TYPE ST_PolarIIChamber_HolderServiceCtrl :
STRUCT
	Gripper : ST_PolarIIChamber_OpenCloseServiceCtrl;
	Rotate : ST_PolarIIChamber_HolderRotateServiceCtrl;
	VacuumEstablish : ST_ServiceCtrl;
END_STRUCT
END_TYPE

(* stored: Version 1.1.0.1, ProductVersion 3.1.4026.18
   DUT ST_PolarIIChamber_HolderServiceCtrl: Id {14000000-0000-0000-0000-000000000064} *)
